(* IEC 61131-3 sources: SortJet_MasterSPS_Aufbau.fbsproj/Device.device.xml.v3^/Plc Logic.plclogic.xml.v3^/Application.application.xml.v3^/00_Basis, 3 files *)

(* ---- Stations_Konfig.gvl ---- *)
(* METADATA
{
	"v3Meta": {
		"objectGuid": "ba3ca572-b5ea-4174-af08-a61d9ddd93e1"
	}
}
*)
{attribute 'allow_unqualified_access'}
NAMESPACE Stations_Konfig
VAR_GLOBAL CONSTANT

//-------------------------------------------------------------------------------------------------
// KONFIG VORHANDENE STATIONEN
//-------------------------------------------------------------------------------------------------

  // Antriebe
  cANZAHL_ANTRIEBE                     : WORD := 29;

  // Ampeln / Hupen
  cANZAHL_AMPELN                       : WORD := 3;
  cANZAHL_HUPEN                        : WORD := 3;

  //Station
  cERSTE_STATION                       : WORD := 201;
  cLETZTE_STATION                      : WORD := 208;

  // Shuttle
  cERSTES_SHUTTLE                      : WORD := 101;
  cLETZTES_SHUTTLE                     : WORD := 102;

  cERSTES_INPUTSHUTTLE                 : WORD := 101;
  cLETZTES_INPUTSHUTTLE                : WORD := 101;

  cERSTES_OUTPUTSHUTTLE                : WORD := 102;
  cLETZTES_OUTPUTSHUTTLE               : WORD := 102;

  // Transfershuttle
  cERSTES_TRANSFERSHUTTLE              : WORD := 151;
  cLETZTES_TRANSFERSHUTTLE             : WORD := 152;

  // Speicher
  cERSTER_SPEICHER                     : WORD := 1;
  cLETZTER_SPEICHER                    : WORD := 1;

  // Faecherwagen
  cERSTE_FAECHERWAGENSTATIONS_NR       : WORD := 301;
  cLETZTE_FAECHERWAGENSTATIONS_NR      : WORD := 305;

  // Hydraulikstationen (Hydraulikaggregate der Faecherwagenstationen Variante Hydraulik)
  cERSTE_HYDRAULIKSTATIONS_NR          : WORD := 1;
  cLETZTE_HYDRAULIKSTATIONS_NR         : WORD := 1;

  // Fremdanlagen
  cERSTE_FREMDANLAGE                   : WORD := 401;
  cLETZTE_FREMDANLAGE                  : WORD := 401;

  cERSTE_FREMDANLAGE_EINLAUF           : WORD := 501;
  cLETZTE_FREMDANLAGE_EINLAUF          : WORD := 501;

  cERSTE_FREMDANLAGE_AUSLAUF           : WORD := 401;
  cLETZTE_FREMDANLAGE_AUSLAUF          : WORD := 401;

  // Terminal
  cERSTES_TERMINAL                     : WORD := 1;
  cLETZTES_TERMINAL                    : WORD := 4;

  // Automatikkreise
  cANZAHL_AUTOMATIKKREISE              : WORD := 2;
  cERSTER_AUTOMATIKKREIS               : WORD := 1;
  cLETZTER_AUTOMATIKKREIS              : WORD := 2;

  // SystemCheck - Shuttle
  cERSTES_SHUTTLESTATIONENSYSTEMCHECK  : WORD := 101;
  cLETZTES_SHUTTLESTATIONENSYSTEMCHECK : WORD := 102;

  // Sicherheitskreise
  cANZAHL_SICHERHEITSKREISE            : WORD := 4;
  cERSTER_SICHERHEITSKREIS             : WORD := 1;
  cLETZTER_SICHERHEITSKREIS            : WORD := 4;

  // Türen
  cANZAHL_TUEREN                       : WORD := 2;
  cERSTE_TUER                          : WORD := 1;
  cLETZTE_TUER                         : WORD := 2;

  // Durchgänge Klappförderer/Türen in der Station
  cANZAHL_DURCHGANGE                   : WORD := 1;
  cERSTER_DURCHGANG                    : WORD := 1;
  cLETZTER_DURCHGANG                   : WORD := 1;

//-------------------------------------------------------------------------------------------------
// KONFIGURATION
//-------------------------------------------------------------------------------------------------
  (* Hinweis:
     - Positionsüberprüfung aller Shuttles und Doppelfördererstationen,da diese als Shuttles gesehne werden
       => Wichtig: Anzahl ist die Ist-Anzahl - 1 [ Teutoglas: 10 Shuttle - 1 ]
  *)
  cANZAHL_SHUTTLE                      : WORD := 2; // Input-, Outputshuttles
  cANZAHL_TRANSFERSHUTTLE              : WORD := 2; // Transfershuttles
  cANZAHL_SHUTTLESTATIONENSYSTEMCHECK  : WORD := 2;

//-------------------------------------------------------------------------------------------------
// DEFINITIONEN
//-------------------------------------------------------------------------------------------------

  // AUTOMATIKKREISE
  cAUTOMATIKKREIS_1                     : WORD := 1;
  cAUTOMATIKKREIS_2                     : WORD := 2;
  cAUTOMATIKKREIS_3                     : WORD := 3;
  cAUTOMATIKKREIS_4                     : WORD := 4;
  cAUTOMATIKKREIS_5                     : WORD := 5;
  cAUTOMATIKKREIS_6                     : WORD := 6;
  cAUTOMATIKKREIS_TRANSFERSHUTTLE       : WORD := 1;

  // STOPP AUTOMATIKKREISE
  cSTOPP_AUTOMATIKKREIS_1                : WORD := 2#0000000000000001;
  cSTOPP_AUTOMATIKKREIS_2                : WORD := 2#0000000000000010;
  cSTOPP_AUTOMATIKKREIS_1_2              : WORD := 2#0000000000000011;
  cSTOPP_AUTOMATIKKREIS_3                : WORD := 2#0000000000000100;
  cSTOPP_AUTOMATIKKREIS_4                : WORD := 2#0000000000001000;
  cSTOPP_AUTOMATIKKREIS_5                : WORD := 2#0000000000010000;
  cSTOPP_AUTOMATIKKREIS_6                : WORD := 2#0000000000100000;
  cSTOPP_AUTOMATIKKREIS_TRANSFERSHUTTLE  : WORD := 2#0000000000001000;
  cSTOPP_ALLE_AUTOMATIKKREIS             : WORD := 2#0000000000000111;

  // WAENDE
  cWAND_DEFAULT                        : WORD := 0;
  cWAND_1                              : WORD := 2#0000000000000001;
  cWAND_2                              : WORD := 2#0000000000000010;
  cWAND_1_2                            : WORD := 2#0000000000000011;
  cANZAHL_WAENDE                       : WORD := 1;

END_VAR

END_NAMESPACE

(* ---- IO_Konfig_Basisbausteine.gvl ---- *)
(* METADATA
{
	"v3Meta": {
		"objectGuid": "1032b1fd-266d-49f6-8f94-6c1a08687c16"
	}
}
*)
{attribute 'allow_unqualified_access'}
NAMESPACE IO_Konfig_Basisbausteine
VAR_CONFIG

// KONFIGURATION: NETZTEILE \ DRUCKLUFT \ ETC.
// *************************************************************************************************

// *************************************************************************************************

  // Druckluft Wartungseinheiten Shuttle (TODO: Eingaenge aus Schaltplan, Platzhalter %MX1.1 = TRUE = OK)
  StatusAnlage.in_bDruckluft_101_OK                                       AT %MX1.1      : BOOL; // OPTION
  StatusAnlage.in_bDruckluft_102_OK                                       AT %IX114.5    : BOOL; // OPTION

//-------------------------------------------------------------------------------------------------
// KONFIGURATION: AMPEL
//-------------------------------------------------------------------------------------------------

  // Ampel AK1 / 1: Speicher Input +01001
  Globale_Bausteine.Ampel_AK[1,1].out_bAmpelLeuchteBlau                     AT %QX2.4    : BOOL; // IO-L - Faecherwagen bereit zum ausschleusen Ampel blau
  Globale_Bausteine.Ampel_AK[1,1].out_bAmpelLeuchteRot                      AT %QX2.3    : BOOL; // IO-L - Automatikkreis Stoerung Ampel rot
  Globale_Bausteine.Ampel_AK[1,1].out_bAmpelLeuchteGelb                     AT %QX2.2    : BOOL; // IO-L - Automatikkreis Hand Ampel gelb
  Globale_Bausteine.Ampel_AK[1,1].out_bAmpelLeuchteGruen                    AT %QX2.1    : BOOL; // IO-L - Automatikkreis Automatik Ampel gruen
  Globale_Bausteine.Horn_AK[1,1].out_bHorn                                  AT %QX2.0    : BOOL; // IO-L - Automatikkreis Checkroutine laeuft Hupe

  // Ampel AK2 / 1: Speicher Output +01001
  Globale_Bausteine.Ampel_AK[2,1].out_bAmpelLeuchteBlau                     AT %QX3.1    : BOOL; // IO-L - Faecherwagen bereit zum ausschleusen Ampel blau
  Globale_Bausteine.Ampel_AK[2,1].out_bAmpelLeuchteRot                      AT %QX3.0    : BOOL; // IO-L - Automatikkreis Stoerung Ampel rot
  Globale_Bausteine.Ampel_AK[2,1].out_bAmpelLeuchteGelb                     AT %QX2.7    : BOOL; // IO-L - Automatikkreis Hand Ampel gelb
  Globale_Bausteine.Ampel_AK[2,1].out_bAmpelLeuchteGruen                    AT %QX2.6    : BOOL; // IO-L - Automatikkreis Automatik Ampel gruen
  Globale_Bausteine.Horn_AK[2,1].out_bHorn                                  AT %QX2.5    : BOOL; // IO-L - Automatikkreis Checkroutine laeuft Hupe

  // Ampel AK2 / 2: Faecherwagenstation +OP4
  Globale_Bausteine.Ampel_AK[2,2].out_bAmpelLeuchteBlau                     AT %QX8.6    : BOOL; // IO-L - Faecherwagen bereit zum ausschleusen Ampel blau
  Globale_Bausteine.Ampel_AK[2,2].out_bAmpelLeuchteRot                      AT %QX8.5    : BOOL; // IO-L - Automatikkreis Stoerung Ampel rot
  Globale_Bausteine.Ampel_AK[2,2].out_bAmpelLeuchteGelb                     AT %QX8.4    : BOOL; // IO-L - Automatikkreis Hand Ampel gelb
  Globale_Bausteine.Ampel_AK[2,2].out_bAmpelLeuchteGruen                    AT %QX8.3    : BOOL; // IO-L - Automatikkreis Automatik Ampel gruen
  Globale_Bausteine.Horn_AK[2,2].out_bHorn                                  AT %QX8.2    : BOOL; // IO-L - Automatikkreis Checkroutine laeuft Hupe

  // Ampel AK1 / 2: Eintransportlinie +OP1
  Globale_Bausteine.Ampel_AK[1,2].out_bAmpelLeuchteBlau                     AT %MX900.0  : BOOL; // OPTION
  Globale_Bausteine.Ampel_AK[1,2].out_bAmpelLeuchteRot                      AT %QX3.6    : BOOL; // IO-L - Automatikkreis Stoerung Ampel rot
  Globale_Bausteine.Ampel_AK[1,2].out_bAmpelLeuchteGelb                     AT %QX3.5    : BOOL; // IO-L - Automatikkreis Hand Ampel gelb
  Globale_Bausteine.Ampel_AK[1,2].out_bAmpelLeuchteGruen                    AT %QX3.4    : BOOL; // IO-L - Automatikkreis Automatik Ampel gruen
  Globale_Bausteine.Horn_AK[1,2].out_bHorn                                  AT %QX3.3    : BOOL; // IO-L - Automatikkreis Checkroutine laeuft Hupe

  // Ampel AK1 / 3: Eintransportlinie +OP2
  Globale_Bausteine.Ampel_AK[1,3].out_bAmpelLeuchteBlau                     AT %MX900.1  : BOOL; // OPTION
  Globale_Bausteine.Ampel_AK[1,3].out_bAmpelLeuchteRot                      AT %QX4.4    : BOOL; // IO-L - Automatikkreis Stoerung Ampel rot
  Globale_Bausteine.Ampel_AK[1,3].out_bAmpelLeuchteGelb                     AT %QX4.3    : BOOL; // IO-L - Automatikkreis Hand Ampel gelb
  Globale_Bausteine.Ampel_AK[1,3].out_bAmpelLeuchteGruen                    AT %QX4.2    : BOOL; // IO-L - Automatikkreis Automatik Ampel gruen
  Globale_Bausteine.Horn_AK[1,3].out_bHorn                                  AT %QX4.1    : BOOL; // IO-L - Automatikkreis Checkroutine laeuft Hupe

  // Ampel AK2 / 3
  Globale_Bausteine.Ampel_AK[2,3].out_bAmpelLeuchteBlau                     AT %MX900.2  : BOOL; // OPTION
  Globale_Bausteine.Ampel_AK[2,3].out_bAmpelLeuchteRot                      AT %MX900.3  : BOOL; // OPTION
  Globale_Bausteine.Ampel_AK[2,3].out_bAmpelLeuchteGelb                     AT %MX900.4  : BOOL; // OPTION
  Globale_Bausteine.Ampel_AK[2,3].out_bAmpelLeuchteGruen                    AT %MX900.5  : BOOL; // OPTION
  Globale_Bausteine.Horn_AK[2,3].out_bHorn                                  AT %MX900.6  : BOOL; // OPTION

//-------------------------------------------------------------------------------------------------
// KONFIGURATION: NETZTEILE \ DRUCKLUFT \ ETC.
//-------------------------------------------------------------------------------------------------

  // HARDWARE EINGAENGE
  StatusAnlage.in_bCAB2_LS_Netzteil_24V_OK                 AT %IX0.4   : BOOL; // IO-L - Netzteil 24V OK
  StatusAnlage.in_bCAB2_KlimaGeraet_OK                     AT %IX0.2   : BOOL; // IO-L - Kuehlgeraet OK
  StatusAnlage.in_bCAB2_LS_Netzfilter_400V_OK              AT %IX0.0   : BOOL; // IO-L - Versorgung 400V Anlage OK
  StatusAnlage.in_bCAB2_LS_400V_OK                         AT %MX1.1   : BOOL; // OPTION
  StatusAnlage.in_bCAB2_LS_24V_Schaltschrank_OK            AT %IX0.5   : BOOL; // IO-L - Sicherungen 24V OK Sammelmeldung Steuerstromkreise Schaltschrank
  StatusAnlage.in_bCAB2_LS_24V_Boxen_OK                    AT %IX0.6   : BOOL; // IO-L - Sicherungen 24V OK Sammelmeldung Steuerstromkreise Anlage
  StatusAnlage.in_bCAB2_LS_230V_OK                         AT %IX0.3   : BOOL; // IO-L - Versorgung OP/PC OK
  StatusAnlage.in_bCAB2_Sicherheitsrelais_201_Kippen_OK    AT %IX3.0   : BOOL; // IO-L - Sicherheitsrelais 201 Hydraulik / kippen OK

END_VAR

END_NAMESPACE

(* ---- StationBasisZuweisungen.prg.st ---- *)
(* METADATA
{
	"v3Meta": {
		"objectGuid": "2c76242e-df1a-45ee-a644-3bee45d641cc"
	}
}
*)
PROGRAM StationBasisZuweisungen
VAR

  // BOOL
  blErsterZyklus              : BOOL := TRUE;

  // WORD
  wlIndex   : WORD;

END_VAR
//-------------------------------------------------------------------------------------------------
// INITIALISIERUNG
//-------------------------------------------------------------------------------------------------
IF ( blErsterZyklus ) THEN

  M_AufrufeZuweisungen();

  // Fehlerinformationen zuweisen
  FOR wlIndex := cERSTE_FAECHERWAGENSTATIONS_NR TO cLETZTE_FAECHERWAGENSTATIONS_NR DO
    IF __ISVALIDREF(starrFaecherwagenBasisParameter[wlIndex].stMKs) THEN
      starrFaecherwagenBasisParameter[wlIndex].awFehlerInformationen[0] := starrFaecherwagenBasisParameter[wlIndex].stMKs.stStationsNummern.NummerExtern;
    END_IF
  END_FOR

  FOR wlIndex := cERSTE_STATION TO cLETZTE_STATION DO
    IF __ISVALIDREF(starrStationBasisParameter[wlIndex].stMKs) THEN
      starrStationBasisParameter[wlIndex].awFehlerInformationen[0] := starrStationBasisParameter[wlIndex].stMKs.stStationsNummern.NummerExtern;
    END_IF
  END_FOR

  FOR wlIndex := cERSTES_SHUTTLE TO cLETZTES_SHUTTLE DO
    IF __ISVALIDREF(starrShuttleBasisParameter[wlIndex].stMKs) THEN
      starrShuttleBasisParameter[wlIndex].awFehlerInformationen[0] := starrShuttleBasisParameter[wlIndex].stMKs.stStationsNummern.NummerExtern;
    END_IF
  END_FOR

  FOR wlIndex := cERSTES_TRANSFERSHUTTLE TO cLETZTES_TRANSFERSHUTTLE DO
    IF __ISVALIDREF(starrTransfershuttleBasisParameter[wlIndex].stMKs) THEN
      starrTransfershuttleBasisParameter[wlIndex].awFehlerInformationen[0] := starrTransfershuttleBasisParameter[wlIndex].stMKs.stStationsNummern.NummerExtern;
    END_IF
  END_FOR

  FOR wlIndex := cERSTE_FREMDANLAGE_AUSLAUF TO cLETZTE_FREMDANLAGE_AUSLAUF DO
    IF __ISVALIDREF(starrFremdanlageAuslaufStationBasisParameter[wlIndex].stMKs) THEN
      starrFremdanlageAuslaufStationBasisParameter[wlIndex].awFehlerInformationen[0] := starrFremdanlageAuslaufStationBasisParameter[wlIndex].stMKs.stStationsNummern.NummerExtern;
    END_IF
  END_FOR

  FOR wlIndex := cERSTE_FREMDANLAGE_EINLAUF TO cLETZTE_FREMDANLAGE_EINLAUF DO
    IF __ISVALIDREF(starrFremdanlageEinlaufStationBasisParameter[wlIndex].stMKs) THEN
      starrFremdanlageEinlaufStationBasisParameter[wlIndex].awFehlerInformationen[0] := starrFremdanlageEinlaufStationBasisParameter[wlIndex].stMKs.stStationsNummern.NummerExtern;
    END_IF
  END_FOR

  blErsterZyklus := FALSE;
END_IF
END_PROGRAM
